(*
SPDX-FileCopyrightText: © 2026 Oleksandr Tiutyk <trofimich@gmail.com>
SPDX-License-Identifier: MIT
License: https://opensource.org/license/mit
*)

(*!
<summary>Names the phases of a filesystem integration regression.</summary>
*)
{attribute 'qualified_only'}
{attribute 'strict'}
TYPE FILE_BUFFER_TEST_PHASE :
(
	//! <summary>prepare directory.</summary>
	PREPARE_DIRECTORY,
	//! <summary>create file.</summary>
	CREATE_FILE,
	//! <summary>wait for file.</summary>
	WAIT_FOR_FILE,
	//! <summary>start invalid operation.</summary>
	START_INVALID_OPERATION,
	//! <summary>wait for invalid operation.</summary>
	WAIT_FOR_INVALID_OPERATION,
	//! <summary>cleanup.</summary>
	CLEANUP
);
END_TYPE

(* stored: Version 1.1.0.1
   DUT FILE_BUFFER_TEST_PHASE: Id {dd49bddf-b5fe-498e-a7aa-48713dc8a2b9} *)
